FUNCTION_BLOCK FB 1
TITLE = A function block without declarations
BEGIN
NETWORK
TITLE = Works on absolute addresses only
      A     I 1.0
      AN    I 1.1
      =     Q 1.0
      L     MW 100
      T     QW 4
END_FUNCTION_BLOCK
